// TIA Portal V20 export
DATA_BLOCK "T5_Resultado"   // DB42901
{ S7_Optimized_Access := 'TRUE' }
AUTHOR : IA
FAMILY : PRUEBA
VERSION : 0.1
// Tanda 1b: un Bool por prueba
// stored: AutoNumber false
   VAR
      L_Inc : Bool;   // Inc
      L_Dec : Bool;   // Dec
      L_MIN : Bool;   // MIN
      L_MAX : Bool;   // MAX
      L_LIMIT : Bool;   // LIMIT
      L_Expt : Bool;   // Expt
      L_DECO : Bool;   // DECO
      L_ENCO : Bool;   // ENCO
      L_SEL : Bool;   // SEL
      L_InRange : Bool;   // IN_RANGE (InRange)
      L_OutRange : Bool;   // OUT_RANGE (OutRange)
      L_OK_NOK : Bool;   // OK / NOT_OK (NOK)
      L_R_TRIG : Bool;   // R_TRIG (DB de instancia T5_Rt_L)
      L_F_TRIG : Bool;   // F_TRIG (DB de instancia T5_Ft_L)
      L_RS : Bool;   // Biestable RS (S_RS)
      L_SET_BF : Bool;   // SET_BF (S_BitfieldCoil)
      L_RESET_BF : Bool;   // [DEDUCIDA] RESET_BF (R_BitfieldCoil)
      L_MOVE_BLK : Bool;   // MOVE_BLK (MoveBlockI)
      L_UMOVE_BLK : Bool;   // UMOVE_BLK (MoveBlockU)
      L_FILL_BLK : Bool;   // FILL_BLK (FillBlockI)
      L_UFILL_BLK : Bool;   // [DEDUCIDA] UFILL_BLK (FillBlockU)
      L_MOVE_BLK_VARIANT : Bool;   // MOVE_BLK_VARIANT
      L_NORM_X : Bool;   // NORM_X (Normalize)
      L_SCALE_X : Bool;   // SCALE_X (Scale_X)
      Vida : DInt;   // Sube cada ciclo
      OK : Int;   // Correctas
      Total : Int := 24;   // Pruebas
      Todo_OK : Bool;   // Todas correctas
   END_VAR
BEGIN
END_DATA_BLOCK
